// TIA Portal V21 export
// export: Created 2026-08-21T20:18:53.5341584Z, ExportSetting None, DisplayName Totally Integrated Automation Portal, DisplayVersion V21, DisplayName STEP 7 Professional, DisplayVersion V21, DisplayName STEP 7 Safety, DisplayVersion V21, DisplayName Tech WebApplication, DisplayVersion V21, DisplayName WinCC Basic/Comfort/Advanced, DisplayVersion V21, DisplayName WinCC Professional, DisplayVersion V21, DisplayName WinCC Unified, DisplayVersion V21
FUNCTION "Flow_Sim" : Void   // FC14, FBD
{ S7_Optimized_Access := 'TRUE' }
// stored: SetENOAutomatically false
   VAR_TEMP
      State : "Service_States";
   END_VAR
BEGIN

REGION Network 1: flow value
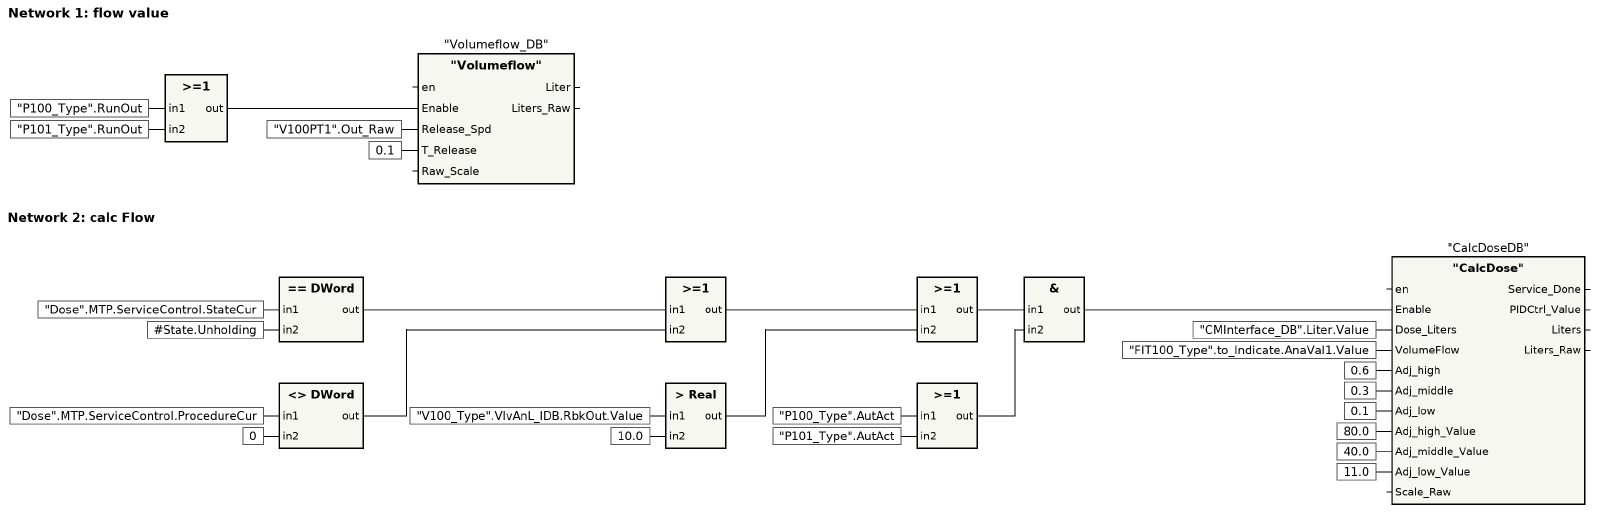
   "Volumeflow_DB"(Enable := "P100_Type".RunOut OR "P101_Type".RunOut,   // "Volumeflow"
                   Release_Spd := "V100PT1".Out_Raw,
                   T_Release := 0.1);
END_REGION

REGION Network 2: calc Flow
   "CalcDoseDB"(Enable := (("Dose".MTP.ServiceControl.StateCur = #State.Unholding) OR ("Dose".MTP.ServiceControl.ProcedureCur <> 0) OR ("V100_Type".VlvAnL_IDB.RbkOut.Value > 10.0)) AND ("P100_Type".AutAct OR "P101_Type".AutAct),   // "CalcDose"
                Dose_Liters := "CMInterface_DB".Liter.Value,
                VolumeFlow := "FIT100_Type".to_Indicate.AnaVal1.Value,
                Adj_high := 0.6,
                Adj_middle := 0.3,
                Adj_low := 0.1,
                Adj_high_Value := 80.0,
                Adj_middle_Value := 40.0,
                Adj_low_Value := 11.0);
END_REGION
END_FUNCTION
